(* IEC 61131-3 sources: repolevel_ST_code_completion/ground_truth/repoeval_Interation_HowTo/readful_result, 2 files *)

(* ---- FirstPublish.st ---- *)
It seems you are working with a repository that involves MQTT communication in Codesys. Based on the provided code fragments, here is a summary of the functionality and structure:

### **Overview of the Code**
1. **MQTT Publisher (`FirstPublish`)**:
   - The `FirstPublish` function block is responsible for publishing messages to an MQTT topic.
   - It initializes an MQTT publisher (`MQTT.MQTTPublish`) and sets the topic (`TestTopic/FromCodesys`) and payload (`testPayload`).
   - The payload is sent when the `doPublish` variable is set to `TRUE`.
   - The `QoS` (Quality of Service) level is set to `ExactlyOnce`, ensuring the message is delivered exactly once.

2. **MQTT Subscriber (`FirstSubscription`)**:
   - The `FirstSubscription` function block subscribes to the same MQTT topic (`TestTopic/FromCodesys`).
   - It uses an MQTT subscription instance (`MQTT.MQTTSubscribe`) and a callback collector (`MQTT.CallbackCollector`) to handle incoming messages.
   - The subscriber is initialized only once (`init` variable ensures this).
   - The `receiver` instance (`MQTT.ReceiveString`) is configured to process messages from the specified topic.

3. **Main Program (`HowTo`)**:
   - The `HowTo` program ties together the publisher and subscriber function blocks.
   - It initializes the MQTT client (`MQTT_IN_OUT`) with the broker URL (`test.mosquitto.org:1883`) and other parameters like timeout and TLS settings.
   - The `FirstPublish` and `FirstSubscription` function blocks are executed in the program.

---

### **Key Features**
1. **MQTT Communication**:
   - The code establishes MQTT communication using the `MQTT_IN_OUT` instance.
   - It connects to the broker (`test.mosquitto.org`) and handles publishing and subscribing.

2. **Topic and Payload**:
   - The topic used for both publishing and subscribing is `TestTopic/FromCodesys`.
   - The payload for publishing is a string (`testPayload`).

3. **Quality of Service (QoS)**:
   - Both publishing and subscribing use `QoS.ExactlyOnce`, ensuring reliable message delivery.

4. **Initialization**:
   - Both function blocks (`FirstPublish` and `FirstSubscription`) use an `init` flag to ensure initialization happens only once.

---

### **Suggestions for Improvement**
1. **Error Handling**:
   - Add error handling for MQTT connection issues, such as broker unavailability or timeout errors.

2. **Dynamic Configuration**:
   - Allow dynamic configuration of the topic, payload, and broker URL instead of hardcoding them.

3. **Logging**:
   - Implement logging to track published and received messages for debugging purposes.

4. **Security**:
   - Consider enabling TLS (`TLS:= TRUE`) for secure communication with the MQTT broker.

---

### **Code Example for Dynamic Configuration**
You could modify the `FirstPublish` and `FirstSubscription` blocks to accept dynamic inputs for the topic and payload:

```st
FUNCTION_BLOCK FirstPublish
VAR_INPUT
    Topic: STRING;
    Payload: STRING;
END_VAR
VAR_OUTPUT
END_VAR
VAR
    publisher: MQTT.MQTTPublish;
    doPublish: BOOL;
    init: BOOL;
END_VAR

IF NOT init THEN
    init := TRUE;
    publisher.SetMqttInOut(MQTT_IN_OUT:= HowTo.MQTT_IN_OUT);
END_IF

publisher(
    Topic:= ADR(Topic),
    PayloadString:= ADR(Payload),
    PublishAsString:= TRUE,
    QoSIn:= MQTT.QoS.ExactlyOnce,
    MRetain:= FALSE,
    send:= doPublish);
```

Similarly, update `FirstSubscription` to accept dynamic inputs for the topic.

---

Let me know if you need further assistance with this code!

(* ---- FirstPublish_1.st ---- *)
It seems you are working with a repository that involves MQTT communication in Codesys. Based on the provided code fragments, here is a summary of the functionality and structure:

### **Overview of the Code**
1. **MQTT Publisher (`FirstPublish`)**:
   - The `FirstPublish` function block is responsible for publishing messages to an MQTT topic.
   - It initializes an MQTT publisher (`MQTT.MQTTPublish`) and sets the topic (`TestTopic/FromCodesys`) and payload (`testPayload`).
   - The payload is sent when the `doPublish` variable is set to `TRUE`.
   - The `QoS` (Quality of Service) level is set to `ExactlyOnce`, ensuring the message is delivered exactly once.

2. **MQTT Subscriber (`FirstSubscription`)**:
   - The `FirstSubscription` function block subscribes to the same MQTT topic (`TestTopic/FromCodesys`).
   - It uses an MQTT subscription instance (`MQTT.MQTTSubscribe`) and a callback collector (`MQTT.CallbackCollector`) to handle incoming messages.
   - The subscriber is initialized only once (`init` variable ensures this).
   - The `receiver` instance (`MQTT.ReceiveString`) is configured to process messages from the specified topic.

3. **Main Program (`HowTo`)**:
   - The `HowTo` program ties together the publisher and subscriber function blocks.
   - It initializes the MQTT client (`MQTT_IN_OUT`) with the broker URL (`test.mosquitto.org:1883`) and other parameters like timeout and TLS settings.
   - The `FirstPublish` and `FirstSubscription` function blocks are executed in the program.

---

### **Key Features**
1. **MQTT Communication**:
   - The code establishes MQTT communication using the `MQTT_IN_OUT` instance.
   - It connects to the broker (`test.mosquitto.org`) and handles publishing and subscribing.

2. **Topic and Payload**:
   - The topic used for both publishing and subscribing is `TestTopic/FromCodesys`.
   - The payload for publishing is a string (`testPayload`).

3. **Quality of Service (QoS)**:
   - Both publishing and subscribing use `QoS.ExactlyOnce`, ensuring reliable message delivery.

4. **Initialization**:
   - Both function blocks (`FirstPublish` and `FirstSubscription`) use an `init` flag to ensure initialization happens only once.

---

### **Suggestions for Improvement**
1. **Error Handling**:
   - Add error handling for MQTT connection issues, such as broker unavailability or timeout errors.

2. **Dynamic Configuration**:
   - Allow dynamic configuration of the topic, payload, and broker URL instead of hardcoding them.

3. **Logging**:
   - Implement logging to track published and received messages for debugging purposes.

4. **Security**:
   - Consider enabling TLS (`TLS:= TRUE`) for secure communication with the MQTT broker.

---

### **Code Example for Dynamic Configuration**
You could modify the `FirstPublish` and `FirstSubscription` blocks to accept dynamic inputs for the topic and payload:

```st
FUNCTION_BLOCK FirstPublish
VAR_INPUT
    Topic: STRING;
    Payload: STRING;
END_VAR
VAR_OUTPUT
END_VAR
VAR
    publisher: MQTT.MQTTPublish;
    doPublish: BOOL;
    init: BOOL;
END_VAR

IF NOT init THEN
    init := TRUE;
    publisher.SetMqttInOut(MQTT_IN_OUT:= HowTo.MQTT_IN_OUT);
END_IF

publisher(
    Topic:= ADR(Topic),
    PayloadString:= ADR(Payload),
    PublishAsString:= TRUE,
    QoSIn:= MQTT.QoS.ExactlyOnce,
    MRetain:= FALSE,
    send:= doPublish);
```

Similarly, update `FirstSubscription` to accept dynamic inputs for the topic.

---

Let me know if you need further assistance with this code!
